(* IEC 61131-3 sources: llm-plc-st-eval/data/processed_definitivo/gpt-4o-2024-08-06/B7/few_shot, 3 files *)

(* ---- ejec_1.st ---- *)
FUNCTION SelBomba : BOOL
VAR_INPUT
    modoAuto : BOOL;   (* Modo automático *)
    btnManual : BOOL;  (* Botón manual *)
    nivelBajo : BOOL;  (* Sensor de nivel bajo *)
END_VAR

(* Selección de la fuente de mando de la bomba *)
(* En modo automático, la bomba enciende si nivelBajo está activo *)
(* En modo manual, la bomba sigue el estado del botón manual *)
SelBomba := (modoAuto AND nivelBajo) OR (NOT modoAuto AND btnManual);
END_FUNCTION

(* ---- ejec_2.st ---- *)
FUNCTION SelBomba : BOOL
VAR_INPUT
    modoAuto : BOOL;    (* Modo automático *)
    btnManual : BOOL;   (* Botón manual *)
    nivelBajo : BOOL;   (* Sensor de nivel bajo *)
END_VAR

(* Selección de la fuente de mando de la bomba *)
IF modoAuto THEN
    SelBomba := nivelBajo; (* En modo automático, la bomba sigue el sensor de nivel bajo *)
ELSE
    SelBomba := btnManual; (* En modo manual, la bomba sigue el botón manual *)
END_IF;
END_FUNCTION

(* ---- ejec_3.st ---- *)
FUNCTION SelBomba : BOOL
VAR_INPUT
    modoAuto : BOOL;   (* Modo automático *)
    btnManual : BOOL;  (* Botón manual *)
    nivelBajo : BOOL;  (* Sensor de nivel bajo *)
END_VAR

(* Selección de la fuente de mando de la bomba *)
IF modoAuto THEN
    (* Modo automático: la bomba enciende si el nivel es bajo *)
    SelBomba := nivelBajo;
ELSE
    (* Modo manual: la bomba sigue el estado del botón manual *)
    SelBomba := btnManual;
END_IF;
END_FUNCTION
